(*
SPDX-FileCopyrightText: © 2026 Oleksandr Tiutyk <trofimich@gmail.com>
SPDX-License-Identifier: MIT
License: https://opensource.org/license/mit
*)

(*
Verifies storage identity, independent snapshot ownership and replacement from a borrowed view.

Keeps the source and predicate instances alive in the owning test task. Teardown clears both predicates
after a successful or failed run.
*)

{attribute 'no_assign'}
{attribute 'no_explicit_call' := 'do not call this function block directly'}
FUNCTION_BLOCK ComparisonPredicateContractsTest EXTENDS TOF_Testing.SingleCycleTest
VAR_STAT
	// Class name shared by instances of this test.
	{attribute 'hide'}
	_ClassName : STRING := __POUNAME();
END_VAR
VAR
	_Source : STRING(24);
	_Storage : TOF_Comparison.SameStoragePredicate;
	_Snapshot : TOF_Comparison.BytewiseEqualityPredicate;
END_VAR

(*
Checks matching text in disjoint storage and the result of mutating the borrowed source.

Replaces the snapshot through its own view, then checks that an enum descriptor with an unsupported
byte size is rejected and leaves the snapshot readable.
*)
METHOD PROTECTED ExecuteTest
VAR
	matchingText : STRING(8) := 'sample';
	sourceValue : __SYSTEM.AnyType;
	query : __SYSTEM.AnyType;
	view : __SYSTEM.AnyType;
	invalidValue : __SYSTEM.AnyType;
	exceptionCode : __SYSTEM.ExceptionCode;
	caught : TOF_Core.IException;
	notSupported : TOF_Core.INotSupportedException;
END_VAR
_Source := matchingText;
sourceValue := TOF_Core.SystemAnyTypes.CreateAnyTypeByAny(anyValue := _Source);
query := TOF_Core.SystemAnyTypes.CreateAnyTypeByAny(anyValue := matchingText);
_Storage.SetReferenceValueByAny(referenceValue := _Source);
_Snapshot.SetReferenceValueByAny(referenceValue := _Source);

Assert.ThatBool(
	actual := _Storage.Check(valueToCompare := sourceValue),
	message := "Storage predicate must accept the original address"
).IsTrue();
Assert.ThatBool(
	actual := _Storage.Check(valueToCompare := query),
	message := "Equal text in a different buffer must fail storage identity"
).IsFalse();
Assert.ThatBool(
	actual := _Snapshot.Check(valueToCompare := query),
	message := "Equal terminated text must match across different capacities"
).IsTrue();

_Source := 'changed';
Assert.ThatBool(
	actual := _Storage.Check(valueToCompare := sourceValue),
	message := "Replacing source content must preserve storage identity"
).IsTrue();
Assert.ThatBool(
	actual := _Snapshot.Check(valueToCompare := sourceValue),
	message := "Replacing source content must leave the owned snapshot independent"
).IsFalse();

view := _Snapshot.ReferenceValue.AsAnyType();
_Snapshot.SetReferenceValueByAnyType(referenceValue := view);
Assert.ThatBool(
	actual := _Snapshot.Check(valueToCompare := query),
	message := "Replacing the owned snapshot from its own view must preserve its text"
).IsTrue();

// Three readable bytes cannot be mapped as an enum by the descriptor factory.
invalidValue.TypeClass := __SYSTEM.TYPE_CLASS.TYPE_ENUM;
invalidValue.pValue := sourceValue.pValue;
invalidValue.diSize := 3;

__TRY
	_Snapshot.SetReferenceValueByAnyType(referenceValue := invalidValue);
__CATCH(exceptionCode)
	caught := TOF_Core.ExceptionManager.GetLastException(
		exceptionCode := exceptionCode,
		catchPointNamespaceName := NamespaceName,
		catchPointPOUName := __POUNAME(),
		catchPointPosition := __POSITION()
	);
__ENDTRY

Assert.ThatBool(
	actual := __QUERYINTERFACE(caught, notSupported),
	message := "Unsupported enum metadata must fail during replacement"
).IsTrue();
Assert.ThatBool(
	actual := _Snapshot.Check(valueToCompare := query),
	message := "Rejected replacement must leave the previous snapshot readable"
).IsTrue();
END_METHOD

(* Clears the borrowed source and releases the owned snapshot for another run. *)
METHOD PROTECTED OnAfterTest
VAR
	emptyValue : __SYSTEM.AnyType;
END_VAR
emptyValue.TypeClass := __SYSTEM.TYPE_CLASS.TYPE_NONE;
emptyValue.pValue := 0;
emptyValue.diSize := 0;
_Storage.SetReferenceValueByAnyType(referenceValue := emptyValue);
_Snapshot.SetReferenceValueByAnyType(referenceValue := emptyValue);
Assert.ThatBool(
	actual := _Storage.ReferenceValue.IsNull AND_THEN _Snapshot.ReferenceValue.IsNull,
	message := "Teardown must clear both predicate descriptors"
).IsTrue();
END_METHOD

// Borrows the concrete class name. Callers must not modify it.
{attribute 'monitoring' := 'call'}
PROPERTY ClassName : REFERENCE TO STRING
GET
ClassName REF= _ClassName;
END_GET
END_PROPERTY

// Borrows the compiler-initialized namespace name. Callers must not modify it.
{attribute 'monitoring' := 'call'}
PROPERTY NamespaceName : REFERENCE TO STRING
GET
NamespaceName REF= CurrentNamespace.Name;
END_GET
END_PROPERTY

// Reports the concrete instance size in bytes.
{attribute 'monitoring' := 'call'}
PROPERTY SelfSize : ULINT
GET
SelfSize := XSIZEOF(THIS^);
END_GET
END_PROPERTY

END_FUNCTION_BLOCK

(* stored: Version 1.1.0.1
   POU ComparisonPredicateContractsTest: Id {389cafd1-13fa-467b-b6a6-251a9ffddd86}, SpecialFunc None
   Method ExecuteTest: Id {eb6c5aeb-5c0e-4e8d-aafb-012686226155}
   Method OnAfterTest: Id {03f0e113-d77f-4be3-a724-03bc9a307220}
   Property ClassName: Id {0be5ca0d-9f50-4774-9233-779f77cc137c}
   Get Get: Id {c2283abc-9e83-4d0d-b5cb-329965ff653e}
   Property NamespaceName: Id {d4ad1406-a17a-4504-9084-f8ee9dc91a65}
   Get Get: Id {72b9d180-0a6b-4a05-8bf5-76b2c5bd0b88}
   Property SelfSize: Id {498f8297-d715-43c7-8fa5-e97a03a7d114}
   Get Get: Id {6eb18f04-6351-4d93-b988-a566bc196cab} *)
